Fanuc KAREL source: KA00154.KL

PROGRAM KA00154
%NOLOCKGROUP
VAR
  SRC: ARRAY[4] OF REAL
  DST: ARRAY[4] OF INTEGER
BEGIN
  DST = SRC
END KA00154
